Fanuc KAREL source: kd00019.KL

-- PROVISIONAL review KL for V940-1; original PC SHA256 3fa4f5185d330107980304e6946cbbf708c064b07167edf3ba733cfa87bb42a1
-- Incomplete behavior may be omitted. Consult companion uncertainty JSON. Do not deploy.
PROGRAM KD00019
%NOLOCKGROUP
VAR
  I : INTEGER
  J : INTEGER
  B : BOOLEAN
  R : REAL
  S : STRING[80]
-- UNRESOLVED_DECL REC type=001100
BEGIN
  -- V9_ZERO_TABLE_METADATA_HINT layout=0001; no indexed target words; source/name/runtime held
  -- UNRESOLVED_PC offsets 5-16; opcodes 9D,22,32,35
  -- UNRESOLVED_PC offsets 26-48; opcodes 22,32,34,9D,52,22,32,35
  -- UNRESOLVED_PC offsets 58-62; opcodes 7F
END KD00019
